(* IEC 61131-3 sources: garage-sweeper/PLC/src/Core, 11 files *)

(* ---- BodyMotion.st ---- *)
TYPE BodyMotion :
STRUCT
	distanceInM : LREAL;
	headingChangeInRad : LREAL;
END_STRUCT
END_TYPE

(* ---- HardwareError.st ---- *)
TYPE HardwareError :
STRUCT
	isActive : BOOL;
	id : UDINT;
	text : STRING(80);
END_STRUCT
END_TYPE

(* ---- LaserScan.st ---- *)
TYPE LaserScan :
STRUCT
	sequence : UDINT;
	startTimestampInNs : ULINT;
	scanDurationInS : REAL;
	angleMinInRad : REAL;
	angleIncrementInRad : REAL;
	count : UINT;
	rangesInM : ARRAY[0..Constants.MAX_SCAN_POINTS - 1] OF REAL;
END_STRUCT
END_TYPE

(* ---- PlatformKind.st ---- *)
{attribute 'qualified_only'}
{attribute 'strict'}
TYPE PlatformKind :
(
	SIMULATION := 0,
	HARDWARE
);
END_TYPE

(* ---- Pose2D.st ---- *)
TYPE Pose2D :
STRUCT
	x : LREAL;
	y : LREAL;
	thetaInRad : LREAL;
END_STRUCT
END_TYPE

(* ---- Twist.st ---- *)
TYPE Twist :
STRUCT
	forwardSpeedInMPerS : LREAL;
	yawRateInRadPerS : LREAL;
END_STRUCT
END_TYPE

(* ---- Vector3.st ---- *)
TYPE Vector3 :
STRUCT
	x : LREAL;
	y : LREAL;
	z : LREAL;
END_STRUCT
END_TYPE

(* ---- WheelSide.st ---- *)
{attribute 'qualified_only'}
{attribute 'strict'}
TYPE WheelSide :
(
	LEFT := 0,
	RIGHT
);
END_TYPE

(* ---- WheelSpeeds.st ---- *)
TYPE WheelSpeeds :
STRUCT
	leftInRadPerS : LREAL;
	rightInRadPerS : LREAL;
END_STRUCT
END_TYPE

(* ---- Constants.st ---- *)
{attribute 'qualified_only'}
VAR_GLOBAL CONSTANT
	MAX_SCAN_POINTS : UINT := 1024;
	SIMULATOR_PROTOCOL_VERSION : UDINT := 1;
	SIMULATOR_TIMEOUT_IN_CYCLES : UDINT := 20;
	LIDAR_TIMEOUT_IN_MS : TIME := T#400MS;
	SIMULATOR_NOT_CONNECTED_ERROR_ID : UDINT := 1001;
	LIDAR_TIMEOUT_ERROR_ID : UDINT := 2001;
END_VAR

(* ---- Parameters.st ---- *)
{attribute 'qualified_only'}
VAR_GLOBAL PERSISTENT
	platform : PlatformKind := PlatformKind.SIMULATION;
	wheelRadiusInM : LREAL := 0.075;
	trackWidthInM : LREAL := 0.40;
	maxWheelSpeedInRadPerS : LREAL := 8.0;
END_VAR
